ADAPTER lamp_control (* Adapter Interface *)
  (* Standard: 61499-1 *)
  (* Version 0.0, 10/23/2026, macie, Schneider Electric *)
  PACKAGE Main;
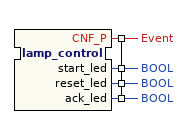
  EVENT_OUTPUT
    CNF_P WITH start_led, reset_led, ack_led; (* Confirmation from Plug *)
  END_EVENT
  VAR_OUTPUT
    start_led : BOOL; (* Confirmation Data from Plug *)
    reset_led : BOOL; (* Indication Data from Plug *)
    ack_led : BOOL;
  END_VAR
  SERVICE SOCKET/PLUG
    SEQUENCE request_confirm
      SOCKET.REQ(REQD) -> PLUG.REQ(REQD);
      PLUG.CNF_P(start_led) -> SOCKET.CNF_P(start_led);
    END_SEQUENCE
    SEQUENCE indication_response
      PLUG.IND(reset_led) -> SOCKET.IND(reset_led);
      SOCKET.RSP(RSPD) -> PLUG.RSP(RSPD);
    END_SEQUENCE
  END_SERVICE
END_ADAPTER
